FUNCTION_BLOCK StartLedControl (* Basic Function Block Type *)
  (* Standard: 61499-2 *)
  (* Version 0.0, 10/21/2026, macie, Schneider Electric, Template *)
  PACKAGE Main;
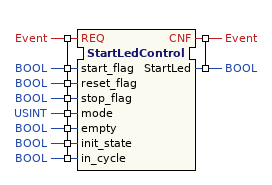
  EVENT_INPUT
    REQ WITH start_flag, reset_flag, stop_flag, mode, empty, init_state, in_cycle; (* Normal Execution Request *)
  END_EVENT
  EVENT_OUTPUT
    CNF WITH StartLed; (* Execution Confirmation *)
  END_EVENT
  VAR_INPUT
    start_flag : BOOL;
    reset_flag : BOOL;
    stop_flag : BOOL; (* Input event qualifier *)
    mode : USINT;
    empty : BOOL;
    init_state : BOOL;
    in_cycle : BOOL;
  END_VAR
  VAR_OUTPUT
    StartLed : BOOL := FALSE; (* Output event qualifier *)
  END_VAR
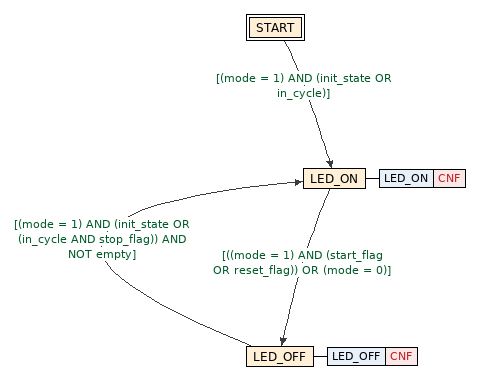
  EC_STATES
    START; (* Initial State *)
    LED_ON : LED_ON -> CNF;
    LED_OFF : LED_OFF -> CNF;
  END_STATES
  EC_TRANSITIONS
    START TO LED_ON := [(mode = 1) AND (init_state OR in_cycle)];
    LED_ON TO LED_OFF := [((mode = 1) AND (start_flag OR reset_flag)) OR (mode = 0)];
    LED_OFF TO LED_ON := [(mode = 1) AND (init_state OR (in_cycle AND stop_flag)) AND NOT empty];
  END_TRANSITIONS
  ALGORITHM LED_ON IN ST:
;
StartLed := TRUE;
  END_ALGORITHM
  ALGORITHM LED_OFF IN ST:
;
StartLed := FALSE;
  END_ALGORITHM
END_FUNCTION_BLOCK
